FUNCTION "ID_Decode_F"   // FC 3, author

VAR_INPUT
   ID : DInt;
END_VAR

VAR_IN_OUT
   ID_Decoded : "ID_Decoded";
END_VAR

VAR_TEMP
   Temp : UInt;
END_VAR

   // RETURN : Void
BEGIN

// Extract XX (first two digits)
#ID_Decoded.Device_Type := #ID / 10000;        // 123456 / 10000 = 12

// Extract YY (middle two digits)
#ID_Decoded.Level := (#ID MOD 10000) / 100; // 123456 % 10000 = 3456 → 3456 / 100 = 34

// Extract ZZ (last two digits)
#ID_Decoded.VTD := #ID MOD 100;       // 123456 % 100 = 56
END_FUNCTION